(* IEC 61131-3 sources: codesys-to-astra/src/POUs/F_C2aWordToHexStr, 2 files *)

(* ---- F_C2aWordToHexStr.decl.st ---- *)
// Назначение: замена OSU.WORD_TO_HEX_STR (OwenStringUtils v3.0, с. 51): WORD -> строка с префиксом и
//             4 hex-символами (дополнение нулями — допущение A9, сверить с ПЛК210), регистр по xUpperCase.
// Автор:      kr0nsch
// Версия:     0.1.0
// Документ:   docs/LIBMAP.md
FUNCTION F_C2aWordToHexStr : STRING(8)
VAR_INPUT
    wInput : WORD;          // исходное значение
    xUpperCase : BOOL;      // TRUE — верхний регистр hex-символов
    sPrefix : STRING(4);    // префикс строки
END_VAR
VAR
    iNibbleNo : INT;        // номер тетрады от старшей
    iNibble : INT;          // значение тетрады 0..15
    sDigits : STRING(16);   // алфавит hex
    sHex : STRING(8);       // hex-часть
END_VAR

(* ---- F_C2aWordToHexStr.impl.st ---- *)
IF xUpperCase THEN
    sDigits := GVL_C2aConst.HEX_DIGITS_UPPER;
ELSE
    sDigits := GVL_C2aConst.HEX_DIGITS_LOWER;
END_IF
sHex := '';
FOR iNibbleNo := GVL_C2aConst.HEX_WORD_DIGITS - 1 TO 0 BY -1 DO
    iNibble := WORD_TO_INT(SHR(wInput, iNibbleNo * GVL_C2aConst.NIBBLE_BITS) AND 16#F);
    sHex := CONCAT(sHex, MID(sDigits, 1, iNibble + 1));
END_FOR
F_C2aWordToHexStr := CONCAT(sPrefix, sHex);
